DATA_BLOCK "S11Recovery"
{ S7_Optimized_Access := 'TRUE' }
VERSION : 0.1
NON_RETAIN
"FB_S11RecoveryRig"
BEGIN
END_DATA_BLOCK
